(* IEC 61131-3 sources: llm-plc-st-eval/data/definitivo/qwen2.5-coder_14b/C6/zero_shot, 1 file *)

(* ---- ejec_1.st ---- *)
1. **Error**: La conversión de `rawTemp` a `tempC` no está realizada correctamente. La fórmula actual divide `rawTemp` por 27648 y luego multiplica por 100, lo que resulta en un valor que no está en el rango de 0.0 a 100.0. La fórmula correcta debería ser `tempC := INT_TO_REAL(rawTemp) / 27648 * 100;`.

2. **Error**: La lógica para controlar el `enfriador` está invertida. El `enfriador` debería activarse cuando `tempC` alcance 80.0 y desactivarse cuando descienda a 75.0. La condición `ELSIF tempC <= 80.0 THEN` debería ser `ELSIF tempC < 75.0 THEN`.

3. **Error**: La lógica para controlar el `enfriador` no conserva su estado entre los umbrales de 75.0 y 80.0. Se necesita una variable de retención para mantener el estado del `enfriador` entre estos umbrales. Se puede agregar una variable interna `enfriadorEstado` para almacenar el estado del `enfriador`.

4. **Error**: La condición para activar `almSensor` cuando `rawTemp` está fuera del rango 0 a 27648 no está completa. También debería considerar el caso cuando `rawTemp` es menor que 0. La condición debería ser `IF rawTemp < 0 OR rawTemp > 27648 THEN`.

**Correcciones propuestas**:

1. **Corrección**: `tempC := INT_TO_REAL(rawTemp) / 27648 * 100;`

2. **Corrección**: `ELSIF tempC < 75.0 THEN`

3. **Corrección**: Agregar una variable interna `enfriadorEstado` y modificar la lógica para controlar el `enfriador`:
    ```pascal
    VAR
        enfriadorEstado : BOOL := FALSE;
    END_VAR

    IF tempC >= 80.0 THEN
        enfriador := TRUE;
        enfriadorEstado := TRUE;
    ELSIF tempC < 75.0 THEN
        enfriador := FALSE;
        enfriadorEstado := FALSE;
    ELSE
        enfriador := enfriadorEstado;
    END_IF
    ```

4. **Corrección**: `IF rawTemp < 0 OR rawTemp > 27648 THEN`
